TYPE T_LintAlias : STRING(80);
END_TYPE

(* stored: Version 1.1.0.1, ProductVersion 3.1.4024.16
   DUT T_LintAlias: Id {3ff34fcb-6ab1-43bd-842c-318285325ff0} *)
